(* IEC 61131-3 sources: codesys-to-astra/tests/POUs/FB_C2aModbus_Test, 6 files *)

(* ---- FB_C2aModbus_Test.decl.st ---- *)
// Назначение: тесты распаковки регистров Modbus REGUL: порядок слов FLOAT32, индекс вне массива, статусы МВ210.
// Автор:      kr0nsch
// Версия:     0.1.0
// Документ:   docs/TEST_REPORT.md
FUNCTION_BLOCK FB_C2aModbus_Test EXTENDS coUnit.FB_TestSuite
VAR CONSTANT
    R_DELTA : REAL := 0.0001;   // допуск сравнения REAL
END_VAR

(* ---- HighWordFirst.method.decl.st ---- *)
// 16#41A0, 16#0000 при HighWordFirst = 20.0 (IEEE 754)
METHOD PRIVATE HighWordFirst
VAR
    rResult : REAL;  // результат
END_VAR

(* ---- LowWordFirst.method.decl.st ---- *)
// 16#0000, 16#41A0 при LowWordFirst = 20.0
METHOD PRIVATE LowWordFirst
VAR
    rResult : REAL;  // результат
END_VAR

(* ---- Mx210Codes.method.decl.st ---- *)
// коды 16#FD, 16#F7 и обычное значение
METHOD PRIVATE Mx210Codes
VAR
    eBreak : E_C2aMx210Status;  // обрыв
    eOff : E_C2aMx210Status;  // отключён
    eOk : E_C2aMx210Status;  // результат
END_VAR

(* ---- UnpackInRange.method.decl.st ---- *)
// FB_C2aMbUnpack: REAL и INT по индексу
METHOD PRIVATE UnpackInRange
VAR
    awData : ARRAY [0..3] OF WORD := [16#C2C8, 16#0000, 16#FFFE, 0];  // -100.0, -2
    fbUnpack : FB_C2aMbUnpack;  // распаковка
END_VAR

(* ---- UnpackOutOfRange.method.decl.st ---- *)
// индекс вне массива -> xValid = FALSE
METHOD PRIVATE UnpackOutOfRange
VAR
    awData : ARRAY [0..1] OF WORD;  // регистры
    fbUnpack : FB_C2aMbUnpack;  // распаковка
END_VAR
